// TIA Portal V20 export
Screen "10_SubMenus"  100x768
  ScreenItem "txtOverview_15" at -2,715 size 100x53  Type=HmiTextBox
  ScreenItem "txtOverview_1" at -2,658 size 100x52  Type=HmiTextBox
  ScreenItem "txtOverview_2" at -2,601 size 100x52  Type=HmiTextBox
  ScreenItem "txtOverview_3" at -2,542 size 100x52  Type=HmiTextBox
  ScreenItem "txtOverview_4" at -2,482 size 100x52  Type=HmiTextBox
  ScreenItem "txtOverview_5" at -2,422 size 100x52  Type=HmiTextBox
  ScreenItem "txtOverview_6" at -2,362 size 100x52  Type=HmiTextBox
  ScreenItem "txtOverview_7" at -2,302 size 100x52  Type=HmiTextBox
  ScreenItem "txtOverview_8" at -2,242 size 100x52  Type=HmiTextBox
  ScreenItem "txtOverview_9" at -2,182 size 100x52  Type=HmiTextBox
  ScreenItem "txtOverview_10" at -2,122 size 100x52  Type=HmiTextBox
  ScreenItem "txtOverview_11" at -2,62 size 100x52  Type=HmiTextBox
  ScreenItem "txtOverview_12" at -2,2 size 100x52  Type=HmiTextBox
  ScreenItem "线_1" at -2,418 size 97x0  Type=HmiLine
